TYPE ST_EL3356ChannelCtrl :
STRUCT
	bStartCalibration			:BOOL;			(* Ctrl start calibration *)
	bDisableCalibration		:BOOL;			(* Ctrl disable calibration *)
	bInputFreeze				:BOOL;			(* Ctrl input freeze *)
	bTare					:BOOL;			(* Ctrl tare *)
END_STRUCT
END_TYPE

(* stored: Version 1.1.0.1, ProductVersion 3.1.4024.15
   DUT ST_EL3356ChannelCtrl: Id {3f428282-8038-4565-9e5e-671712aa3675} *)
